(* IEC 61131-3 sources: llm-plc-st-eval/codesys/dobles/B3, 4 files *)

(* ---- 01_Correcta.st ---- *)
(* DOBLE DE PRUEBA B3/Correcta - NO ES CORPUS. Esperado: veredicto 1 *)
FUNCTION_BLOCK FB_Contador
VAR_INPUT
    sensorPieza : BOOL;
    btnReset : BOOL;
END_VAR
VAR_OUTPUT
    loteListo : BOOL;
    cuenta : INT;
END_VAR
VAR
    prev : BOOL;
END_VAR
IF btnReset THEN
    cuenta := 0;
    loteListo := FALSE;
ELSIF sensorPieza AND NOT prev THEN
    cuenta := cuenta + 1;
END_IF
IF cuenta >= 12 THEN
    loteListo := TRUE;
END_IF
prev := sensorPieza;
END_FUNCTION_BLOCK

(* ---- 02_CuentaPorNivel.st ---- *)
(* DOBLE DE PRUEBA B3/CuentaPorNivel - NO ES CORPUS. Esperado: veredicto 2, falla en el paso 2 *)
FUNCTION_BLOCK FB_Contador
VAR_INPUT
    sensorPieza : BOOL;
    btnReset : BOOL;
END_VAR
VAR_OUTPUT
    loteListo : BOOL;
    cuenta : INT;
END_VAR
VAR
    prev : BOOL;
END_VAR
IF btnReset THEN
    cuenta := 0;
    loteListo := FALSE;
ELSIF sensorPieza THEN
    cuenta := cuenta + 1;
END_IF
IF cuenta >= 12 THEN
    loteListo := TRUE;
END_IF
prev := sensorPieza;
END_FUNCTION_BLOCK

(* ---- 03_PresetIncorrecto.st ---- *)
(* DOBLE DE PRUEBA B3/PresetIncorrecto - NO ES CORPUS. Esperado: veredicto 2, falla en el paso 4 *)
FUNCTION_BLOCK FB_Contador
VAR_INPUT
    sensorPieza : BOOL;
    btnReset : BOOL;
END_VAR
VAR_OUTPUT
    loteListo : BOOL;
    cuenta : INT;
END_VAR
VAR
    prev : BOOL;
END_VAR
IF btnReset THEN
    cuenta := 0;
    loteListo := FALSE;
ELSIF sensorPieza AND NOT prev THEN
    cuenta := cuenta + 1;
END_IF
IF cuenta >= 10 THEN
    loteListo := TRUE;
END_IF
prev := sensorPieza;
END_FUNCTION_BLOCK

(* ---- 04_ResetIncompleto.st ---- *)
(* DOBLE DE PRUEBA B3/ResetIncompleto - NO ES CORPUS. Esperado: veredicto 2, falla en el paso 6 *)
FUNCTION_BLOCK FB_Contador
VAR_INPUT
    sensorPieza : BOOL;
    btnReset : BOOL;
END_VAR
VAR_OUTPUT
    loteListo : BOOL;
    cuenta : INT;
END_VAR
VAR
    prev : BOOL;
END_VAR
IF btnReset THEN
    cuenta := 0;
ELSIF sensorPieza AND NOT prev THEN
    cuenta := cuenta + 1;
END_IF
IF cuenta >= 12 THEN
    loteListo := TRUE;
END_IF
prev := sensorPieza;
END_FUNCTION_BLOCK
